Staubli VAL3: _supervisorTasks.pgx

public program _supervisorTasks()
  local num l_i
  local bool l_bResult
begin
  for l_i = 0 to size(_nClock)-1
    _nClock[l_i]=0
  endFor
  do
    //任务监控
    if taskStatus("plc")>1 and (clock()-_nClock[1]>5)
      _nClock[1]=clock()
      taskResume("plc",0)
      rs:bIsError=true
    else
      _nClock[1]=clock()
    endIf
    if taskStatus("appMain")>1 and (clock()-_nClock[2]>5)
      _nClock[2]=clock()
      rs:bIsError=true
      taskResume("appMain",0)
    else
      _nClock[2]=clock()
    endIf
    if taskStatus("HMI")>1
      //保存当前数据
      bTosave=true
      call trajectory:onSave(bTosave)
      bTosave=true
      call program:onSave(bTosave)
      wait(rs:bIsSaving==false)
      l_bResult=userPageConfirm("需要重载HMI应用？")
      if l_bResult

        taskKill("HMI")
        wait(taskStatus("HMI")==-1)
        taskCreate "HMI",50,home:main()
        wait(taskStatus("HMI")==1)
      endIf
    endIf


    delay(0)
  until false
end
